TYPE ST_UnitReq :
STRUCT
	bPSetActive	: BOOL;
	fPSet		: REAL;		// kW, 유닛 출력
	bQSetActive	: BOOL;
	fQSet		: REAL;		// kvar
END_STRUCT
END_TYPE

(* stored: Version 1.1.0.1, ProductVersion 3.1.4024.15
   DUT ST_UnitReq: Id {76f58a11-46ed-4305-bebf-b1a40d257e79} *)
